// FC_TIME_TO_DINT: TIME转DINT (占位版本)
// 描述: 在LSP环境中返回0, 避免类型转换错误

FUNCTION FC_TIME_TO_DINT : DINT
VAR_INPUT
    TimeValue : TIME;
END_VAR

BEGIN
    // [多平台占位] LSP环境返回0
    // TIA Portal: FC_TIME_TO_DINT := DINT(#TimeValue) / 1000;
    FC_TIME_TO_DINT := 0;

END_FUNCTION
